(* Tests that the base and log-record ProtoJSON serializers write the OTLP/JSON wire form: field encodings, failure reasons, and resource/scope grouping. *)
FUNCTION_BLOCK FB_TestProtoJsonSerializer EXTENDS FB_TestSuite

THIS^.testSerializeNumberValues();
THIS^.testSerializeLogRecord();
THIS^.testSerializeLogRecordWithoutTraceIdOmitsFlags();
THIS^.testSerializeRejectsNullInputs();
THIS^.testSerializeLogsDataGroupsByResourceAndScope();

(* A null log-record pointer or a null member key fails serialization with its own failure reason,
   so a caller can tell a missing record from a serializer misuse instead of writing broken JSON. *)
METHOD testSerializeRejectsNullInputs : REFERENCE TO FB_Test
VAR
	serializer: FB_LogRecordProtoJsonSerializer;
	root: SJsonValue;
	records: SJsonValue;
	pRecord: POINTER TO FB_LogRecord;
	serializationSucceeded: BOOL;
	failureReason: E_ProtoJsonSerializerFailureReason;
END_VAR
TcUnit.TEST('testSerializeRejectsNullInputs');
	root := serializer.parser.NewDocument();
	root := serializer.parser.SetObject(root);
	records := serializer.parser.AddArrayMember(root, 'logRecords', 0);

	// pRecord is deliberately left 0.
	serializationSucceeded := serializer.serializeLogRecord(
		v:=records,
		pLogRecord:=pRecord,
		failureReason=>failureReason
	);
	THIS^.AssertFalse(serializationSucceeded, 'Expected a null log-record pointer to fail serialization');
	THIS^.AssertTrue(
		failureReason = E_ProtoJsonSerializerFailureReason.LOG_RECORD_POINTER_NULL,
		'Expected LOG_RECORD_POINTER_NULL as the failure reason for a null log record'
	);

	// pKey is deliberately 0.
	serializationSucceeded := serializer.serializeUint32Value(
		v:=root,
		pKey:=0,
		val:=1,
		failureReason=>failureReason
	);
	THIS^.AssertFalse(serializationSucceeded, 'Expected a null JSON member key to fail serialization');
	THIS^.AssertTrue(
		failureReason = E_ProtoJsonSerializerFailureReason.KEY_POINTER_NULL,
		'Expected KEY_POINTER_NULL as the failure reason for a null member key'
	);
TcUnit.TEST_FINISHED();
END_METHOD

(* A record built through the logger serializes every field in its OTLP/JSON form: enums and fixed32 as numbers,
   64-bit integers as decimal strings, trace and span IDs as hex, and values as typed AnyValue objects. *)
METHOD testSerializeLogRecord : REFERENCE TO FB_Test
VAR
	resource: FB_Resource(schemaUrl:='');
	provider: FB_LoggerProvider(resource:=resource);
	scope: FB_InstrumentationScope(name:='motor1', version:='0.0.1a', schemaUrl:='');
	logger: FB_Logger(scope:=scope, provider:=provider);
	processor: FB_LogRecordProcessor_ForRecordInspection(0);
	serializer: FB_LogRecordProtoJsonSerializer();
	emitSuccess: BOOL;
	emitFailureResult: E_LoggerFailureReason;
	timestamp: ULINT := 1581452773000000789;
	traceId: ARRAY [0..15] OF BYTE := [0, 1, 2, 3, 4, 5, 6, 7, 8, 9, 10, 11, 12, 13, 14, 15];
	spanId: ARRAY [0..7] OF BYTE := [16, 17, 18, 19, 20, 21, 22, 23];
	durationMs: DINT := 42;
	temperature: LREAL := 21.5;
	pRecord: POINTER TO FB_LogRecord;
	root: SJsonValue;
	records: SJsonValue;
	obj: SJsonValue;
	member: SJsonValue;
	attributes: SJsonValue;
	attribute: SJsonValue;
	value: SJsonValue;
	actualString: STRING;
	serializationSucceeded: BOOL;
	serializerFailureReason: E_ProtoJsonSerializerFailureReason;
END_VAR
TcUnit.TEST('testSerializeLogRecord');
	processor.free();
	logger.free();

	// Create a representative record through the public logger API.
	logger
		.startLogRecord(severityNumber:=E_SeverityNumber.DEBUG)
		.setTimestamp(timestamp)
		.setEventName('Serialization Event')
		.setBody('This is a body string value')
		._setTraceId(ADR(traceId), SIZEOF(traceId))
		._setSpanId(ADR(spanId), SIZEOF(spanId))
		._setFlags(16#01)  // sampled
		.setStringAttribute('stats.label', 'pVal')
		.setNumberAttribute('stats.duration_ms', durationMs)
		.setNumberAttribute('stats.temperature', temperature);
	THIS^.AssertTrue(logger.pLogRecord <> 0, 'Expected the logger to hold a log record before emission');
	IF logger.pLogRecord <> 0 THEN
		// no builder sets droppedAttributesCount; set by hand to check it is written
		logger.pLogRecord^.droppedAttributesCount := 2;
	END_IF

	emitSuccess := logger.emit(failureResult=>emitFailureResult);
	THIS^.AssertTrue(emitSuccess, 'Expected log record emission to succeed');
	provider
		.stageProcessor(processor)
		.tick();
	THIS^.AssertTrue(processor.lastOperationSucceeded, 'Expected the inspection processor to capture the emitted record');
	THIS^.AssertTrue(logger.pLogRecord = 0, 'Expected emit to release the logger-owned record');
	pRecord := processor.pop();
	THIS^.AssertTrue(pRecord <> 0, 'Expected the processor to return the emitted record');
	IF pRecord <> 0 THEN

	// serializeLogRecord appends one LogRecord object to the supplied JSON array.
	root := serializer.parser.NewDocument();
	serializer.parser.SetObject(root);
	records := serializer.parser.AddArrayMember(root, 'logRecords', 0);
	serializationSucceeded := serializer.serializeLogRecord(
		v:=records,
		pLogRecord:=pRecord,
		failureReason=>serializerFailureReason
	);
	THIS^.AssertTrue(
		serializationSucceeded AND_THEN serializerFailureReason = E_ProtoJsonSerializerFailureReason.NA,
		'Expected LogRecord serialization to succeed without a failure reason'
	);
	obj := serializer.parser.GetArrayValueByIdx(records, 0);
		THIS^.AssertTrue(serializer.parser.IsObject(obj), 'Expected the logRecords array to hold one LogRecord object');

		// OTLP/JSON encodes enums and fixed32 values as numbers.
		// 5 is DEBUG; flags 1 is the sampled trace flag of the record's span.
		member := serializer.parser.FindMember(obj, 'severityNumber');
		THIS^.AssertEquals_UDINT(5, serializer.parser.GetUint(member), 'Expected severityNumber 5 (DEBUG) as a JSON number');
		actualString := serializer.parser.GetString(serializer.parser.FindMember(obj, 'severityText'));
		THIS^.AssertEquals_STRING('DEBUG', actualString, 'Expected severityText to be the severity enum name');
		THIS^.AssertEquals_UDINT(1, serializer.parser.GetUint(serializer.parser.FindMember(obj, 'flags')), 'Expected flags 1 (sampled) as a JSON number');
		THIS^.AssertEquals_UDINT(2, serializer.parser.GetUint(serializer.parser.FindMember(obj, 'droppedAttributesCount')), 'Expected droppedAttributesCount 2 as a JSON number');

		// OTLP/JSON encodes 64-bit integers as decimal strings and trace/span IDs as hex.
		actualString := serializer.parser.GetString(serializer.parser.FindMember(obj, 'timeUnixNano'));
		THIS^.AssertEquals_STRING('1581452773000000789', actualString, 'Expected string-encoded timeUnixNano');
		actualString := serializer.parser.GetString(serializer.parser.FindMember(obj, 'traceId'));
		THIS^.AssertEquals_STRING('000102030405060708090A0B0C0D0E0F', actualString, 'Expected hex-encoded traceId');
		actualString := serializer.parser.GetString(serializer.parser.FindMember(obj, 'spanId'));
		THIS^.AssertEquals_STRING('1011121314151617', actualString, 'Expected hex-encoded spanId');

		// Event name and body.
		actualString := serializer.parser.GetString(serializer.parser.FindMember(obj, 'eventName'));
		THIS^.AssertEquals_STRING('Serialization Event', actualString, 'Expected eventName to be written as set');
		value := serializer.parser.FindMember(serializer.parser.FindMember(obj, 'body'), 'stringValue');
		actualString := serializer.parser.GetString(value);
		THIS^.AssertEquals_STRING('This is a body string value', actualString, 'Expected AnyValue string body');

		// Attributes keep insertion order; each value is a typed AnyValue, with intValue as a decimal string.
		attributes := serializer.parser.FindMember(obj, 'attributes');
		THIS^.AssertTrue(serializer.parser.IsArray(attributes), 'Expected attributes to be a JSON array');
		attribute := serializer.parser.GetArrayValueByIdx(attributes, 0);
		actualString := serializer.parser.GetString(serializer.parser.FindMember(attribute, 'key'));
		THIS^.AssertEquals_STRING('stats.label', actualString, 'Expected string attribute key');
		value := serializer.parser.FindMember(serializer.parser.FindMember(attribute, 'value'), 'stringValue');
		actualString := serializer.parser.GetString(value);
		THIS^.AssertEquals_STRING('pVal', actualString, 'Expected string attribute AnyValue');
		attribute := serializer.parser.GetArrayValueByIdx(attributes, 1);
		actualString := serializer.parser.GetString(serializer.parser.FindMember(attribute, 'key'));
		THIS^.AssertEquals_STRING('stats.duration_ms', actualString, 'Expected numeric attribute key');
		value := serializer.parser.FindMember(serializer.parser.FindMember(attribute, 'value'), 'intValue');
		actualString := serializer.parser.GetString(value);
		THIS^.AssertEquals_STRING('42', actualString, 'Expected numeric attribute AnyValue');
		attribute := serializer.parser.GetArrayValueByIdx(attributes, 2);
		actualString := serializer.parser.GetString(serializer.parser.FindMember(attribute, 'key'));
		THIS^.AssertEquals_STRING('stats.temperature', actualString, 'Expected floating attribute key');
		value := serializer.parser.FindMember(serializer.parser.FindMember(attribute, 'value'), 'doubleValue');
		THIS^.AssertTrue(serializer.parser.IsDouble(value) AND_THEN serializer.parser.GetDouble(value) = 21.5, 'Expected floating attribute AnyValue');
	END_IF

	IF pRecord <> 0 THEN pRecord^.delete(pSelf:=pRecord); END_IF
	processor.free();
	logger.free();

TcUnit.TEST_FINISHED();
END_METHOD

(* A record without a trace id belongs to no trace, so the serializer leaves out flags even when the record holds some,
   along with traceId and spanId. The record stores flags as set; omitting them is the serializer's decision. *)
METHOD testSerializeLogRecordWithoutTraceIdOmitsFlags : REFERENCE TO FB_Test
VAR
	resource: FB_Resource(schemaUrl:='');
	provider: FB_LoggerProvider(resource:=resource);
	scope: FB_InstrumentationScope(name:='motor1', version:='0.0.1a', schemaUrl:='');
	logger: FB_Logger(scope:=scope, provider:=provider);
	processor: FB_LogRecordProcessor_ForRecordInspection(0);
	serializer: FB_LogRecordProtoJsonSerializer();
	emitSuccess: BOOL;
	emitFailureResult: E_LoggerFailureReason;
	pRecord: POINTER TO FB_LogRecord;
	root: SJsonValue;
	records: SJsonValue;
	obj: SJsonValue;
	serializationSucceeded: BOOL;
	serializerFailureReason: E_ProtoJsonSerializerFailureReason;
END_VAR
TcUnit.TEST('testSerializeLogRecordWithoutTraceIdOmitsFlags');
	emitSuccess := logger
		.startLogRecord(severityNumber:=E_SeverityNumber.INFO)
		._setFlags(16#01)  // sampled, but no trace id
		.emit(failureResult=>emitFailureResult);
	THIS^.AssertTrue(emitSuccess, 'Expected log record emission to succeed');
	provider
		.stageProcessor(processor)
		.tick();
	pRecord := processor.pop();
	THIS^.AssertTrue(pRecord <> 0, 'Expected the processor to return the emitted record');
	IF pRecord <> 0 THEN
		THIS^.AssertEquals_UDINT(1, pRecord^.flags, 'Expected the record to keep the flags it was given');

		root := serializer.parser.NewDocument();
		serializer.parser.SetObject(root);
		records := serializer.parser.AddArrayMember(root, 'logRecords', 0);
		serializationSucceeded := serializer.serializeLogRecord(
			v:=records,
			pLogRecord:=pRecord,
			failureReason=>serializerFailureReason
		);
		THIS^.AssertTrue(serializationSucceeded, 'Expected LogRecord serialization to succeed');
		obj := serializer.parser.GetArrayValueByIdx(records, 0);
		THIS^.AssertTrue(serializer.parser.IsObject(obj), 'Expected the logRecords array to hold one LogRecord object');
		THIS^.AssertTrue(serializer.parser.FindMember(obj, 'flags') = 0, 'Expected no flags member without a trace id');
		THIS^.AssertTrue(serializer.parser.FindMember(obj, 'traceId') = 0, 'Expected no traceId member');
		THIS^.AssertTrue(serializer.parser.FindMember(obj, 'spanId') = 0, 'Expected no spanId member');
		pRecord^.delete(pSelf:=pRecord);
	END_IF
	processor.free();
TcUnit.TEST_FINISHED();
END_METHOD

(* serializeLogsData groups interleaved records into one ResourceLogs per resource and one ScopeLogs per scope,
   in first-seen order with records kept in arrival order, and drains the queue it is given. *)
METHOD testSerializeLogsDataGroupsByResourceAndScope : REFERENCE TO FB_Test
VAR
	resourceB: FB_Resource('resource.b');
	resourceA: FB_Resource('resource.a');
	resourceC: FB_Resource('resource.c');
	providerB: FB_LoggerProvider(resource:=resourceB);
	providerA: FB_LoggerProvider(resource:=resourceA);
	providerC: FB_LoggerProvider(resource:=resourceC);
	scopeB: FB_InstrumentationScope('scope.b', '1.0.0', 'scope.b.schema');
	scopeA: FB_InstrumentationScope('scope.a', '1.0.0', 'scope.a.schema');
	scopeC: FB_InstrumentationScope('scope.c', '1.0.0', 'scope.c.schema');
	loggerBb: FB_Logger(scope:=scopeB, provider:=providerB);
	loggerBa: FB_Logger(scope:=scopeA, provider:=providerB);
	loggerAc: FB_Logger(scope:=scopeC, provider:=providerA);
	loggerAb: FB_Logger(scope:=scopeB, provider:=providerA);
	loggerCa: FB_Logger(scope:=scopeA, provider:=providerC);
	processor: FB_LogRecordProcessor_ForRecordsInspection(
		maxQueueSize:=0,
		scheduledDelayMillis:=1000,
		maxExportBatchSize:=512,
		exporter:=0
	);
	queue: REFERENCE TO FB_LogRecordQueue;
	serializer: FB_LogRecordProtoJsonSerializer;
	emitSucceeded: BOOL;
	_idx: UDINT;
	resourceLogs: SJsonValue;
	resourceObj: SJsonValue;
	scopeLogs: SJsonValue;
	scopeObj: SJsonValue;
	logRecords: SJsonValue;
	recordObj: SJsonValue;
	actualString: STRING;
	serializationSucceeded: BOOL;
	serializerFailureReason: E_ProtoJsonSerializerFailureReason;
END_VAR
TcUnit.TEST('testSerializeLogsDataGroupsByResourceAndScope');
	processor.free();
	queue REF= processor.records;

	// ---- Arrange: eight records with interleaved resource/scope pairs ----
	// Each logger is one resource/scope pair, named resource then scope (loggerBa is resource B, scope A).
	// The timestamp is the record number, so each record can be identified in the output.
	//   record:   1  2  3  4  5  6  7  8
	//   resource: B  A  C  B  C  A  B  A
	//   scope:    B  C  A  A  A  B  B  C
	FOR _idx := 1 TO 8 DO
		CASE _idx OF
			1, 7: emitSucceeded := THIS^._emitRecord(logger:=loggerBb, provider:=providerB, processor:=processor, timestamp:=_idx);
			4:    emitSucceeded := THIS^._emitRecord(logger:=loggerBa, provider:=providerB, processor:=processor, timestamp:=_idx);
			2, 8: emitSucceeded := THIS^._emitRecord(logger:=loggerAc, provider:=providerA, processor:=processor, timestamp:=_idx);
			6:    emitSucceeded := THIS^._emitRecord(logger:=loggerAb, provider:=providerA, processor:=processor, timestamp:=_idx);
			3, 5: emitSucceeded := THIS^._emitRecord(logger:=loggerCa, provider:=providerC, processor:=processor, timestamp:=_idx);
		END_CASE
		THIS^.AssertTrue(emitSucceeded, CONCAT('Expected record ', CONCAT(UDINT_TO_STRING(_idx), ' to reach the processor')));
	END_FOR
	THIS^.AssertEquals_UDINT(8, queue.count, 'Expected eight records queued before serialization');

	// ---- Act ----
	serializationSucceeded := serializer.serializeLogsData(
		logRecords:=queue,
		failureReason=>serializerFailureReason
	);
	THIS^.AssertTrue(
		serializationSucceeded AND_THEN serializerFailureReason = E_ProtoJsonSerializerFailureReason.NA,
		'Expected LogsData serialization to succeed without a failure reason'
	);
	THIS^.AssertEquals_UDINT(0, queue.count, 'Expected the serializer to drain the queue it was given');

	// ---- Assert: three ResourceLogs groups in first-seen order B, A, C ----
	resourceLogs := serializer.parser.FindMember(serializer.jsonValue, 'resourceLogs');
	THIS^.AssertTrue(resourceLogs <> 0 AND_THEN serializer.parser.IsArray(resourceLogs), 'Expected resourceLogs to be a JSON array');

	THIS^.AssertTrue(serializer.parser.GetArrayValueByIdx(resourceLogs, 3) = 0, 'Expected exactly three ResourceLogs groups');

	// Resource B was seen first. Its scope B records remain in arrival order,
	// followed by the later first-seen scope A group.
	resourceObj := serializer.parser.GetArrayValueByIdx(resourceLogs, 0);
	actualString := serializer.parser.GetString(serializer.parser.FindMember(resourceObj, 'schemaUrl'));
	THIS^.AssertEquals_STRING('resource.b', actualString, 'Expected resource B as the first ResourceLogs group');
	scopeLogs := serializer.parser.FindMember(resourceObj, 'scopeLogs');
	scopeObj := serializer.parser.GetArrayValueByIdx(scopeLogs, 0);

	actualString := serializer.parser.GetString(serializer.parser.FindMember(serializer.parser.FindMember(scopeObj, 'scope'), 'name'));
	THIS^.AssertEquals_STRING('scope.b', actualString, 'Expected scope B as the first scope of resource B');
	logRecords := serializer.parser.FindMember(scopeObj, 'logRecords');
	recordObj := serializer.parser.GetArrayValueByIdx(logRecords, 0);

	actualString := serializer.parser.GetString(serializer.parser.FindMember(recordObj, 'timeUnixNano'));
	THIS^.AssertEquals_STRING('1', actualString, 'Expected record 1 first in resource B scope B');
	recordObj := serializer.parser.GetArrayValueByIdx(logRecords, 1);
	actualString := serializer.parser.GetString(serializer.parser.FindMember(recordObj, 'timeUnixNano'));
	THIS^.AssertEquals_STRING('7', actualString, 'Expected record 7 second in resource B scope B');
	THIS^.AssertTrue(serializer.parser.GetArrayValueByIdx(logRecords, 2) = 0, 'Expected exactly two records in resource B scope B');

	scopeObj := serializer.parser.GetArrayValueByIdx(scopeLogs, 1);
	actualString := serializer.parser.GetString(serializer.parser.FindMember(serializer.parser.FindMember(scopeObj, 'scope'), 'name'));
	THIS^.AssertEquals_STRING('scope.a', actualString, 'Expected scope A as the second scope of resource B');
	logRecords := serializer.parser.FindMember(scopeObj, 'logRecords');
	recordObj := serializer.parser.GetArrayValueByIdx(logRecords, 0);

	actualString := serializer.parser.GetString(serializer.parser.FindMember(recordObj, 'timeUnixNano'));
	THIS^.AssertEquals_STRING('4', actualString, 'Expected record 4 in resource B scope A');
	THIS^.AssertTrue(serializer.parser.GetArrayValueByIdx(logRecords, 1) = 0, 'Expected exactly one record in resource B scope A');
	THIS^.AssertTrue(serializer.parser.GetArrayValueByIdx(scopeLogs, 2) = 0, 'Expected exactly two scopes for resource B');

	// Resource A was seen second. Its repeated scope C records are one group.
	resourceObj := serializer.parser.GetArrayValueByIdx(resourceLogs, 1);
	actualString := serializer.parser.GetString(serializer.parser.FindMember(resourceObj, 'schemaUrl'));
	THIS^.AssertEquals_STRING('resource.a', actualString, 'Expected resource A as the second ResourceLogs group');
	scopeLogs := serializer.parser.FindMember(resourceObj, 'scopeLogs');
	scopeObj := serializer.parser.GetArrayValueByIdx(scopeLogs, 0);

	actualString := serializer.parser.GetString(serializer.parser.FindMember(serializer.parser.FindMember(scopeObj, 'scope'), 'name'));
	THIS^.AssertEquals_STRING('scope.c', actualString, 'Expected scope C as the first scope of resource A');
	logRecords := serializer.parser.FindMember(scopeObj, 'logRecords');
	recordObj := serializer.parser.GetArrayValueByIdx(logRecords, 0);

	actualString := serializer.parser.GetString(serializer.parser.FindMember(recordObj, 'timeUnixNano'));
	THIS^.AssertEquals_STRING('2', actualString, 'Expected record 2 first in resource A scope C');
	recordObj := serializer.parser.GetArrayValueByIdx(logRecords, 1);

	actualString := serializer.parser.GetString(serializer.parser.FindMember(recordObj, 'timeUnixNano'));
	THIS^.AssertEquals_STRING('8', actualString, 'Expected record 8 second in resource A scope C');
	THIS^.AssertTrue(serializer.parser.GetArrayValueByIdx(logRecords, 2) = 0, 'Expected exactly two records in resource A scope C');

	scopeObj := serializer.parser.GetArrayValueByIdx(scopeLogs, 1);
	actualString := serializer.parser.GetString(serializer.parser.FindMember(serializer.parser.FindMember(scopeObj, 'scope'), 'name'));
	THIS^.AssertEquals_STRING('scope.b', actualString, 'Expected scope B as the second scope of resource A');
	logRecords := serializer.parser.FindMember(scopeObj, 'logRecords');
	recordObj := serializer.parser.GetArrayValueByIdx(logRecords, 0);
	actualString := serializer.parser.GetString(serializer.parser.FindMember(recordObj, 'timeUnixNano'));
	THIS^.AssertEquals_STRING('6', actualString, 'Expected record 6 in resource A scope B');
	THIS^.AssertTrue(serializer.parser.GetArrayValueByIdx(logRecords, 1) = 0, 'Expected exactly one record in resource A scope B');
	THIS^.AssertTrue(serializer.parser.GetArrayValueByIdx(scopeLogs, 2) = 0, 'Expected exactly two scopes for resource A');

	// Resource C was seen third and its non-adjacent records share one scope.
	resourceObj := serializer.parser.GetArrayValueByIdx(resourceLogs, 2);
	actualString := serializer.parser.GetString(serializer.parser.FindMember(resourceObj, 'schemaUrl'));
	THIS^.AssertEquals_STRING('resource.c', actualString, 'Expected resource C as the third ResourceLogs group');
	scopeLogs := serializer.parser.FindMember(resourceObj, 'scopeLogs');
	scopeObj := serializer.parser.GetArrayValueByIdx(scopeLogs, 0);
	actualString := serializer.parser.GetString(serializer.parser.FindMember(serializer.parser.FindMember(scopeObj, 'scope'), 'name'));
	THIS^.AssertEquals_STRING('scope.a', actualString, 'Expected scope A as the only scope of resource C');
	logRecords := serializer.parser.FindMember(scopeObj, 'logRecords');
	recordObj := serializer.parser.GetArrayValueByIdx(logRecords, 0);
	actualString := serializer.parser.GetString(serializer.parser.FindMember(recordObj, 'timeUnixNano'));
	THIS^.AssertEquals_STRING('3', actualString, 'Expected record 3 first in resource C scope A');
	recordObj := serializer.parser.GetArrayValueByIdx(logRecords, 1);
	actualString := serializer.parser.GetString(serializer.parser.FindMember(recordObj, 'timeUnixNano'));
	THIS^.AssertEquals_STRING('5', actualString, 'Expected record 5 second in resource C scope A');
	THIS^.AssertTrue(serializer.parser.GetArrayValueByIdx(logRecords, 2) = 0, 'Expected exactly two records in resource C scope A');
	THIS^.AssertTrue(serializer.parser.GetArrayValueByIdx(scopeLogs, 1) = 0, 'Expected exactly one scope for resource C');

	processor.free();
TcUnit.TEST_FINISHED();
END_METHOD

(* Integers up to 32 bits and finite floats are written as JSON numbers, while 64-bit integers and
   NaN/Infinity are written as strings, as ProtoJSON requires so that no value loses precision or breaks JSON. *)
METHOD testSerializeNumberValues : REFERENCE TO FB_Test
VAR
	serializer: FB_BaseProtoJsonSerializer;
	root: SJsonValue;
	nSInt: SINT := -12;
	nInt: INT := -1234;
	nDInt: DINT := -123456789;
	nLInt: LINT := -9007199254740993; // -(2^53 + 1): cannot be held exactly by a JSON (double) number
	nUSInt: USINT := 12;
	nUInt: UINT := 1234;
	nUDInt: UDINT := 4000000000;
	nULInt: ULINT := 18000000000000000000; // above 2^63, so it only fits an unsigned 64-bit integer
	fReal: REAL := 42.25;
	fLReal: LREAL := -24.5;
	fNaN: LREAL;
	fPositiveInfinity: LREAL;
	fNegativeInfinity: LREAL;
	// IEEE 754 double bit patterns; ST has no literals for these values.
	nNaNBits: LWORD := LWORD#16#7FF8000000000000;
	nPositiveInfinityBits: LWORD := LWORD#16#7FF0000000000000;
	nNegativeInfinityBits: LWORD := LWORD#16#FFF0000000000000;
	member: SJsonValue;
	actualString: STRING;
END_VAR
TcUnit.TEST('testSerializeNumberValues');
	root := serializer.parser.NewDocument();
	serializer.parser.SetObject(root);

	// serializeNumberValue takes ANY_NUM and dispatches on the actual type.
	THIS^.AssertTrue(serializer.serializeNumberValue(root, ADR('sintValue'), nSInt), 'Expected a SINT to serialize');
	THIS^.AssertTrue(serializer.serializeNumberValue(root, ADR('intValue'), nInt), 'Expected an INT to serialize');
	THIS^.AssertTrue(serializer.serializeNumberValue(root, ADR('dintValue'), nDInt), 'Expected a DINT to serialize');
	THIS^.AssertTrue(serializer.serializeNumberValue(root, ADR('lintValue'), nLInt), 'Expected a LINT to serialize');
	THIS^.AssertTrue(serializer.serializeNumberValue(root, ADR('usintValue'), nUSInt), 'Expected a USINT to serialize');
	THIS^.AssertTrue(serializer.serializeNumberValue(root, ADR('uintValue'), nUInt), 'Expected a UINT to serialize');
	THIS^.AssertTrue(serializer.serializeNumberValue(root, ADR('udintValue'), nUDInt), 'Expected a UDINT to serialize');
	THIS^.AssertTrue(serializer.serializeNumberValue(root, ADR('ulintValue'), nULInt), 'Expected a ULINT to serialize');
	THIS^.AssertTrue(serializer.serializeNumberValue(root, ADR('realValue'), fReal), 'Expected a REAL to serialize');
	THIS^.AssertTrue(serializer.serializeNumberValue(root, ADR('lrealValue'), fLReal), 'Expected an LREAL to serialize');

	THIS^.AssertEquals_DINT(-12, serializer.parser.GetInt(serializer.parser.FindMember(root, 'sintValue')), 'Expected SINT as a JSON number');
	THIS^.AssertEquals_DINT(-1234, serializer.parser.GetInt(serializer.parser.FindMember(root, 'intValue')), 'Expected INT as a JSON number');
	THIS^.AssertEquals_DINT(-123456789, serializer.parser.GetInt(serializer.parser.FindMember(root, 'dintValue')), 'Expected DINT as a JSON number');
	actualString := serializer.parser.GetString(serializer.parser.FindMember(root, 'lintValue'));
	THIS^.AssertEquals_STRING('-9007199254740993', actualString, 'Expected LINT as a decimal JSON string');
	THIS^.AssertEquals_UDINT(12, serializer.parser.GetUint(serializer.parser.FindMember(root, 'usintValue')), 'Expected USINT as a JSON number');
	THIS^.AssertEquals_UDINT(1234, serializer.parser.GetUint(serializer.parser.FindMember(root, 'uintValue')), 'Expected UINT as a JSON number');
	THIS^.AssertEquals_UDINT(4000000000, serializer.parser.GetUint(serializer.parser.FindMember(root, 'udintValue')), 'Expected UDINT as a JSON number');
	actualString := serializer.parser.GetString(serializer.parser.FindMember(root, 'ulintValue'));
	THIS^.AssertEquals_STRING('18000000000000000000', actualString, 'Expected ULINT as a decimal JSON string');
	member := serializer.parser.FindMember(root, 'realValue');
	THIS^.AssertTrue(serializer.parser.IsDouble(member) AND_THEN serializer.parser.GetDouble(member) = 42.25, 'Expected REAL as a JSON number');
	member := serializer.parser.FindMember(root, 'lrealValue');
	THIS^.AssertTrue(serializer.parser.IsDouble(member) AND_THEN serializer.parser.GetDouble(member) = -24.5, 'Expected LREAL as a JSON number');

	// ProtoJSON requires special floating-point values to be quoted strings.
	MEMCPY(ADR(fNaN), ADR(nNaNBits), SIZEOF(fNaN));
	MEMCPY(ADR(fPositiveInfinity), ADR(nPositiveInfinityBits), SIZEOF(fPositiveInfinity));
	MEMCPY(ADR(fNegativeInfinity), ADR(nNegativeInfinityBits), SIZEOF(fNegativeInfinity));
	serializer.serializeNumberValue(root, ADR('nanValue'), fNaN);
	serializer.serializeNumberValue(root, ADR('positiveInfinityValue'), fPositiveInfinity);
	serializer.serializeNumberValue(root, ADR('negativeInfinityValue'), fNegativeInfinity);
	actualString := serializer.parser.GetString(serializer.parser.FindMember(root, 'nanValue'));
	THIS^.AssertEquals_STRING('NaN', actualString, 'Expected NaN as the quoted string NaN');
	actualString := serializer.parser.GetString(serializer.parser.FindMember(root, 'positiveInfinityValue'));
	THIS^.AssertEquals_STRING('Infinity', actualString, 'Expected positive infinity as the quoted string Infinity');
	actualString := serializer.parser.GetString(serializer.parser.FindMember(root, 'negativeInfinityValue'));
	THIS^.AssertEquals_STRING('-Infinity', actualString, 'Expected negative infinity as the quoted string -Infinity');

TcUnit.TEST_FINISHED();
END_METHOD

(*
	Emits one INFO record stamped with timestamp through logger, then ticks its provider with the
	processor staged, so the record reaches the processor now and records keep their emit order
	across providers.
*)
METHOD _emitRecord : BOOL
VAR_INPUT
	logger: REFERENCE TO FB_Logger;
	provider: REFERENCE TO FB_LoggerProvider;
	processor: REFERENCE TO FB_LogRecordProcessor_Base;
	timestamp: ULINT;
END_VAR
VAR
	emitFailureReason: E_LoggerFailureReason;
END_VAR
_emitRecord := logger
	.startLogRecord(severityNumber:=E_SeverityNumber.INFO)
	.setTimestamp(timestamp)
	.emit(failureResult=>emitFailureReason);
_emitRecord := _emitRecord AND_THEN provider
	.stageProcessor(processor)
	.tick();
END_METHOD

END_FUNCTION_BLOCK

(* stored: Version 1.1.0.1
   POU FB_TestProtoJsonSerializer: Id {355aaa54-d854-4f5d-a742-3803c7661c44}, SpecialFunc None
   Method testSerializeRejectsNullInputs: Id {e9865385-1f56-43aa-b979-d2dbed1ed025}
   Method testSerializeLogRecord: Id {432059f0-a68e-4217-85ac-25035b48c8cb}
   Method testSerializeLogRecordWithoutTraceIdOmitsFlags: Id {e1cf92e3-492f-4c8f-9263-cefaa68cf72c}
   Method testSerializeLogsDataGroupsByResourceAndScope: Id {3baae409-f1cd-4ee8-b8e2-c63cbc28a66d}
   Method testSerializeNumberValues: Id {802e0990-b061-4995-9126-6b3d466b4e43}
   Method _emitRecord: Id {8f74556f-15f5-4254-923d-1c6d25a6b693} *)
